FUNCTION_BLOCK AKid_Object EXTENDS TcoCore.TcoObject

END_FUNCTION_BLOCK

(* stored: Version 1.1.0.1, ProductVersion 3.1.4024.6
   POU AKid_Object: Id {212108e8-9c8f-0055-088d-793993f095ba}, SpecialFunc None *)
